// TIA Portal V20 export
TYPE "HMI_Achse_Positionen_überschreiben"
   STRUCT
      Wert_Position_Überschreiben : Array[0..16] of Real;
      Wert_Speed_Überschreiben : Array[0..16] of Real;
      Trig_Position_Überschreiben : Array[0..16] of Bool;
   END_STRUCT;
END_TYPE
